# EPICS substitutions: db/Beckhoff_7XXX/ecmcEX72XX_OPT_touchProbe.substitutions
file "ecmcEL72XX_TP.template"
{
  pattern {CH_ID}
          {"$(OPT_CH_ID=01)"}
}
